Fanuc KAREL source: kd00057.KL

-- PROVISIONAL review KL for V770-1; original PC SHA256 2df413a0de430b58e47245683cfa187a83dd2c1a0f64a08b9d060c2280f7a047
-- Incomplete behavior may be omitted. Consult companion uncertainty JSON. Do not deploy.
PROGRAM KD00057
%NOLOCKGROUP
VAR
  I : INTEGER
  J : INTEGER
  B : BOOLEAN
  R : REAL
  S : STRING[80]
-- UNRESOLVED_DECL P type=000101
-- UNRESOLVED_DECL Q type=000101
BEGIN
  -- UNRESOLVED_PC offsets 5-37; opcodes 01,22,1C,06,22,1C,07,82,0B
  -- UNRESOLVED_PC offsets 42-46; opcodes 7F
END KD00057
